(* IEC 61131-3 sources: PortalRobot/Portal_robot/Device/application/ST/ST_GEOMETRY_CONTROL, 7 files *)

(* ---- ST_GEOMETRY_CALL.st ---- *)
TYPE ST_GEOMETRY_CALL :
STRUCT
	udiId : UDINT; // Не меняется от вызова до результата контроля
	uiMachine : UINT;
	uiProductType : UINT;
	uiStation : UINT; // 0 до автоматического выбора свободного ГК
	xForced : BOOL;
	uiState : UINT; // 1 вызван, 2 в захвате/ожидание, 3 доставка, 4 на ГК, 5 в магазине, 6 отменён, 7 прерван, 8 изъят
	uiReason : UINT; // 1 заняты оба ГК, 2 нет доступного ГК, 3 отключён, 4 авария, 5 перезапуск/неопределённость
	uiMagazine : UINT;
	uiPallet : UINT;
	uiSlot : UINT;
END_STRUCT
END_TYPE

(* ---- ST_GEOMETRY_CONFIG.st ---- *)
TYPE ST_GEOMETRY_CONFIG :
STRUCT
	xConfigured : BOOL;
	lrX : LREAL;
	lrY : LREAL;
	lrZ : LREAL;
	lrSafeZ : LREAL := -300.0; // Signed-смещение безопасного подхода от рабочей Z
	lrChangeZ : LREAL := -150.0; // Legacy-поле OPC UA; маршрут использует SAFE_Z, при записи равно lrSafeZ
	lrSpeedFactor : LREAL := 0.2;
END_STRUCT
END_TYPE

(* ---- ST_GEOMETRY_EVENT.st ---- *)
TYPE ST_GEOMETRY_EVENT :
STRUCT
	udiSequence : UDINT;
	udiTimeMs : UDINT; // Монотонные часы PLC, не настенные часы
	uiEnvironment : UINT; // NORMAL=0, SIMULATION=1, SC500_BENCH=2
	Call : ST_GEOMETRY_CALL;
END_STRUCT
END_TYPE

(* ---- ST_GEOMETRY_MEMORY.st ---- *)
TYPE ST_GEOMETRY_MEMORY :
STRUCT
	xOccupied : BOOL;
	xRecoveryRequired : BOOL;
	xAtEndSeen : BOOL; // Потерю датчика считаем изъятием только после прихода на него
	dwAlarm : DWORD;
	xRobotStopLatched : BOOL;
	udiLastDepositId : UDINT;
	udiProducedPartsTotal : UDINT;
	Part : ST_GEOMETRY_CALL;
END_STRUCT
END_TYPE

(* ---- ST_GEOMETRY_REQUEST.st ---- *)
TYPE ST_GEOMETRY_REQUEST :
STRUCT
	uiAction : UINT; // 1 Enable, 2 Disable, 3 Confirm, 4 Reject, 5 ManualRun, 6 Stop, 7 RemoveSimulation, 8 Call, 9 Auto, 10 Period, 11 Config, 12 Cancel, 13 Capture, 14 SimAlarm, 15 SimAlarmClear, 16 CellSettings
	uiStation : UINT;
	uiMachine : UINT;
	udiValue : UDINT;
	Config : ST_GEOMETRY_CONFIG;
END_STRUCT
END_TYPE

(* ---- ST_GEOMETRY_SIGNALS.st ---- *)
TYPE ST_GEOMETRY_SIGNALS :
STRUCT
	xReserve : BOOL;
	xDeposited : BOOL;
	xReleased : BOOL;
	xRobotInteraction : BOOL;
	Call : ST_GEOMETRY_CALL;
END_STRUCT
END_TYPE

(* ---- ST_GEOMETRY_STATUS.st ---- *)
TYPE ST_GEOMETRY_STATUS :
STRUCT
	uiState : UINT; // 0 выключен, 1 свободен, 2 передача роботом, 3 транспорт, 4 ждёт изъятия, 5 восстановление, 6 авария, 7 ручной ход
	xEnabled : BOOL;
	xReady : BOOL;
	xOccupied : BOOL;
	xPartStored : BOOL; // Подтверждённая укладка, отдельно от резерва и неизвестности
	xReserved : BOOL;
	xPartAtEnd : BOOL;
	xDriveRunning : BOOL;
	xDriveAlarm : BOOL;
	xError : BOOL;
	xRobotStopRequired : BOOL;
	xEnableAllowed : BOOL;
	xDisableAllowed : BOOL;
	xConfirmAllowed : BOOL;
	xConfirmationActive : BOOL;
	xRecoveryRequired : BOOL; // Проверка всей ленты нужна независимо от попытки включения
	xManualStartAllowed : BOOL;
	xResetAllowed : BOOL;
	xResetBusy : BOOL;
	xConfigAllowed : BOOL;
	xPointWriteAllowed : BOOL; // Запись данных: связь/SoftMotion/валидные лимиты, без технологических блокировок
	xSimulationRemoveAllowed : BOOL;
	xSimulationAlarmAllowed : BOOL;
	xConfigured : BOOL;
	udiProducedPartsTotal : UDINT;
	udiPartId : UDINT;
	uiMachine : UINT;
	uiProductType : UINT;
	rTravel : REAL; // Положение модели 0..1; в NORMAL только оценка для изображения
	dwEnableBlockers : DWORD; // Причины запрета команды включения; 0 = xEnableAllowed
	dwConfirmBlockers : DWORD; // Причины запрета подтверждения пустоты; 0 = xConfirmAllowed
	xCallWaitWarning : BOOL; // Активный W52 ячейки; снимается подтверждением предупреждений
	xDisablePending : BOOL; // Штатное выключение ждёт завершения доставки и останова ленты
END_STRUCT
END_TYPE
